FUNCTION_BLOCK TcoDigitalInspectorTests EXTENDS TcoInspectorTests
VAR
    _sut            : TcoInspectors.TcoDigitalInspector(THIS^);
    _inspectedValue : BOOL;
END_VAR

METHOD Inspect : TcoInspectors.IInspector
Inspect := _sut.Inspect(_inspectedValue);
END_METHOD

METHOD PROTECTED Main
SUPER^.Main();
END_METHOD

METHOD  WithCoordinator : REFERENCE TO TcoInspectorTests
VAR_INPUT
	inoCoordinator : TcoCore.ITcoCoordinator;
END_VAR
_sut.WithCoordinator(_coordinator);
WithCoordinator REF= THIS^;
END_METHOD

END_FUNCTION_BLOCK

(* stored: Version 1.1.0.1, ProductVersion 3.1.4024.9
   POU TcoDigitalInspectorTests: Id {006ccc7b-92fd-0f72-19d8-beb7c19c5ae1}, SpecialFunc None
   Method Inspect: Id {3859c7f2-f312-0dbb-12dd-249af68ea862}
   Method Main: Id {0585db86-c979-0f41-16cb-a6ae8111e25a}
   Method WithCoordinator: Id {40f16ac7-8430-09d1-0ef0-083e86fb63ad} *)
